FUNCTION_BLOCK SortingCommandFrame (* Sorting-only architecture following Distribution and tutorial modules 1-4 *)
  (* Standard: 61499-2 *)
  (* Version 2.0, 2026-11-09, sorting2n, sorting2n *)
  PACKAGE Main;
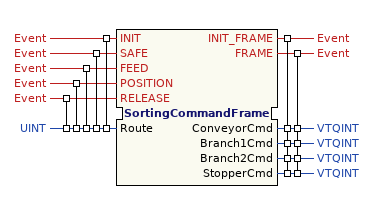
  EVENT_INPUT
    INIT WITH Route;
    SAFE WITH Route;
    FEED WITH Route;
    POSITION WITH Route;
    RELEASE WITH Route;
  END_EVENT
  EVENT_OUTPUT
    INIT_FRAME WITH ConveyorCmd, Branch1Cmd, Branch2Cmd, StopperCmd;
    FRAME WITH ConveyorCmd, Branch1Cmd, Branch2Cmd, StopperCmd;
  END_EVENT
  VAR_INPUT
    Route : UINT := 0;
  END_VAR
  VAR_OUTPUT
    ConveyorCmd : VTQINT;
    Branch1Cmd : VTQINT;
    Branch2Cmd : VTQINT;
    StopperCmd : VTQINT;
  END_VAR
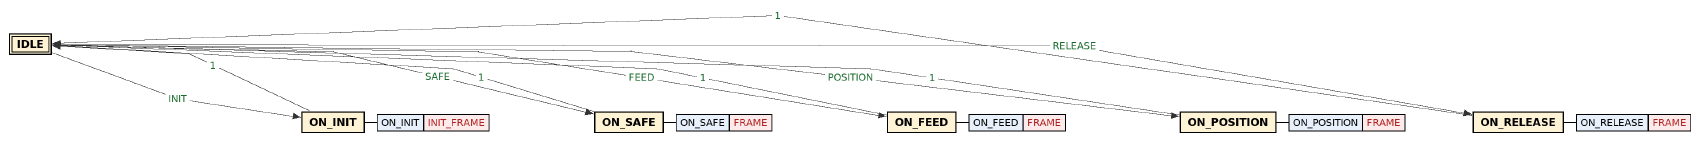
  EC_STATES
    IDLE;
    ON_INIT : ON_INIT -> INIT_FRAME;
    ON_SAFE : ON_SAFE -> FRAME;
    ON_FEED : ON_FEED -> FRAME;
    ON_POSITION : ON_POSITION -> FRAME;
    ON_RELEASE : ON_RELEASE -> FRAME;
  END_STATES
  EC_TRANSITIONS
    IDLE TO ON_INIT := INIT;
    ON_INIT TO IDLE := 1;
    IDLE TO ON_SAFE := SAFE;
    ON_SAFE TO IDLE := 1;
    IDLE TO ON_FEED := FEED;
    ON_FEED TO IDLE := 1;
    IDLE TO ON_POSITION := POSITION;
    ON_POSITION TO IDLE := 1;
    IDLE TO ON_RELEASE := RELEASE;
    ON_RELEASE TO IDLE := 1;
  END_TRANSITIONS
  ALGORITHM ON_INIT IN ST:
ConveyorCmd.value := 2; ConveyorCmd.quality := 0;
Branch1Cmd.value := 2; Branch1Cmd.quality := 0;
Branch2Cmd.value := 2; Branch2Cmd.quality := 0;
StopperCmd.value := 0; StopperCmd.quality := 0;
  END_ALGORITHM
  ALGORITHM ON_SAFE IN ST:
ConveyorCmd.value := 2; ConveyorCmd.quality := 0;
Branch1Cmd.value := 2; Branch1Cmd.quality := 0;
Branch2Cmd.value := 2; Branch2Cmd.quality := 0;
StopperCmd.value := 0; StopperCmd.quality := 0;
  END_ALGORITHM
  ALGORITHM ON_FEED IN ST:
ConveyorCmd.value := 1; ConveyorCmd.quality := 0;
Branch1Cmd.value := 2; Branch1Cmd.quality := 0;
Branch2Cmd.value := 2; Branch2Cmd.quality := 0;
StopperCmd.value := 0; StopperCmd.quality := 0;
  END_ALGORITHM
  ALGORITHM ON_POSITION IN ST:
ConveyorCmd.value := 1; ConveyorCmd.quality := 0;
Branch1Cmd.value := 2; Branch1Cmd.quality := 0;
Branch2Cmd.value := 2; Branch2Cmd.quality := 0;
StopperCmd.value := 0; StopperCmd.quality := 0;
IF Route = 1 THEN Branch1Cmd.value := 1; ELSIF Route = 2 THEN Branch2Cmd.value := 1; END_IF;
  END_ALGORITHM
  ALGORITHM ON_RELEASE IN ST:
ConveyorCmd.value := 1; ConveyorCmd.quality := 0;
Branch1Cmd.value := 2; Branch1Cmd.quality := 0;
Branch2Cmd.value := 2; Branch2Cmd.quality := 0;
StopperCmd.value := 1; StopperCmd.quality := 0;
IF Route = 1 THEN Branch1Cmd.value := 1; ELSIF Route = 2 THEN Branch2Cmd.value := 1; END_IF;
  END_ALGORITHM
END_FUNCTION_BLOCK
